Universal Robots PolyScope program: krc_tending.urp

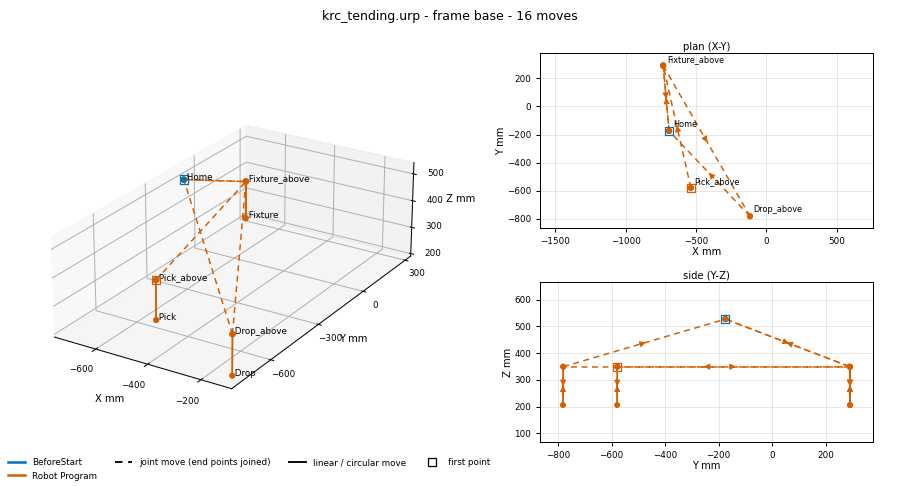
[picture p0: tool path of krc_tending.urp in frame base, 16 of 17 moves have a stored position in this frame; points joined in program order, loops and branches not executed]
Program krc_tending (installation=krc_cell directory=/programs createdIn=5.12.7.1102192 lastSavedIn=5.12.7.1102192 robotSerialNumber=20195299999)
Calibrated DH parameters: a=[0, -0.6127, -0.57155, 0, 0, 0]; d=[0.1807, 0, 0, 0.17415, 0.11985, 0.11655]; alpha=[1.570796, 0, 0, 1.570796, -1.570796, 0]; deltaTheta=[0, 0, 0, 0, 0, 0]
InitVariablesNode
BeforeStart
  'First move: to where the arm already is, so starting the program never moves it on its own'
  start_pose := get_actual_tcp_pose()
  MoveL speed 150 mm/s, acceleration 500 mm/s^2 (useActiveTCP=true optimoveEnabled=false optiMoveSpeed=0.3 optiMoveAcceleration=0.09) feature=Base
    Waypoint Start_pose (Variable): variable=start_pose
  'Every start: clear the handshake, then check it's at home before it moves at all'
  Set ExpressionOutput pin=GP_int_out[5]; expression=10
  Set ExpressionOutput pin=GP_int_out[1]; expression=0
  Set ExpressionOutput pin=GP_int_out[2]; expression=0
  Set ExpressionOutput pin=GP_int_out[3]; expression=0
  Set ExpressionOutput pin=GP_int_out[4]; expression=0
  beat := 0
  home_q := [0.0, -1.57, 1.57, -1.57, -1.57, 0.0]
  q_now := get_actual_joint_positions()
  If norm(q_now[0]-home_q[0])>0.05 or norm(q_now[1]-home_q[1])>0.05 or norm(q_now[2]-home_q[2])>0.05 or norm(q_now[3]-home_q[3])>0.05 or norm(q_now[4]-home_q[4])>0.05 or norm(q_now[5]-home_q[5])>0.05
    'Stopped mid-move last time: moving home from here could hit the fixture or the part, so it doesn't try'
    Set ExpressionOutput pin=GP_int_out[5]; expression=900
    Popup Error (haltProgram=true message=The robot is away from home. Jog it home, then press Start on the panel. inputType=Text)
  Set DigitalOutput pin=tool_out[0]; digitalValue=0
  Wait Sleep waitTime=0.5
  MoveJ speed 57.3 deg/s, acceleration 68.75 deg/s^2 (useActiveTCP=true optimoveEnabled=false optiMoveSpeed=0.3 optiMoveAcceleration=0.09) feature=Base
    Waypoint Home: TCP in base x=-691.676 y=-174.362 z=526.755 mm, rx=2.2206 ry=2.2206 rz=0 rad; joints [0, -89.954, 89.954, -89.954, -89.954, 0] deg; TCP offset x=0 y=0 z=150 mm, rx=0 ry=0 rz=0 rad
Robot Program (runOnlyOnce=false)
  Folder Ready
    'At home, waiting for a command'
    Set ExpressionOutput pin=GP_int_out[5]; expression=100
    Set ExpressionOutput pin=GP_int_out[1]; expression=1
    Wait Condition expression=GP_int_in[1]≟1 or GP_int_in[1]≟2
  Folder Acknowledge
    'Echo the command, and stop being ready while busy'
    cmd := GP_int_in[1]
    Set ExpressionOutput pin=GP_int_out[1]; expression=0
    Set ExpressionOutput pin=GP_int_out[2]; expression=cmd
    ok := True
  If cmd≟1
    'Load: pick a part from the tray, place it in the fixture'
    Set ExpressionOutput pin=GP_int_out[5]; expression=200
    MoveJ speed 57.3 deg/s, acceleration 68.75 deg/s^2 (useActiveTCP=true optimoveEnabled=false optiMoveSpeed=0.3 optiMoveAcceleration=0.09) feature=Base
      Waypoint Pick_above: TCP in base x=-536.89 y=-578.569 z=348.935 mm, rx=2.2208 ry=2.2208 rz=0.001 rad; joints [34.377, -80.214, 97.403, -107.143, -89.954, 34.377] deg
    MoveL speed 150 mm/s, acceleration 500 mm/s^2 (useActiveTCP=true optimoveEnabled=false optiMoveSpeed=0.3 optiMoveAcceleration=0.09) feature=Base
      Waypoint Pick: TCP in base x=-537.712 y=-579.131 z=205.685 mm, rx=2.2208 ry=2.2208 rz=0.001 rad; joints [34.377, -74.485, 105.997, -121.467, -89.954, 34.377] deg
    Set DigitalOutput pin=tool_out[0]; digitalValue=1
    Wait Sleep waitTime=0.5
    MoveL speed 150 mm/s, acceleration 500 mm/s^2 (useActiveTCP=true optimoveEnabled=false optiMoveSpeed=0.3 optiMoveAcceleration=0.09) feature=Base
      Waypoint Pick_above: TCP in base x=-536.89 y=-578.569 z=348.935 mm, rx=2.2208 ry=2.2208 rz=0.001 rad; joints [34.377, -80.214, 97.403, -107.143, -89.954, 34.377] deg
    If tool_out[0]≟False
      'Gripper missed the part'
      ok := False
    Else 
      MoveJ speed 57.3 deg/s, acceleration 68.75 deg/s^2 (useActiveTCP=true optimoveEnabled=false optiMoveSpeed=0.3 optiMoveAcceleration=0.09) feature=Base
        Waypoint Fixture_above: TCP in base x=-733.795 y=290.754 z=348.935 mm, rx=2.2208 ry=2.2208 rz=-0.001 rad; joints [-34.377, -80.214, 97.403, -107.143, -89.954, -34.377] deg
      Set ExpressionOutput pin=GP_int_out[5]; expression=210
      Wait Condition expression=GP_int_in[2]≟1
      MoveL speed 150 mm/s, acceleration 500 mm/s^2 (useActiveTCP=true optimoveEnabled=false optiMoveSpeed=0.3 optiMoveAcceleration=0.09) feature=Base
        Waypoint Fixture: TCP in base x=-734.617 y=291.316 z=205.685 mm, rx=2.2208 ry=2.2208 rz=-0.001 rad; joints [-34.377, -74.485, 105.997, -121.467, -89.954, -34.377] deg
      Set ExpressionOutput pin=GP_int_out[5]; expression=220
      Set DigitalOutput pin=tool_out[0]; digitalValue=0
      Wait Sleep waitTime=0.5
      MoveL speed 150 mm/s, acceleration 500 mm/s^2 (useActiveTCP=true optimoveEnabled=false optiMoveSpeed=0.3 optiMoveAcceleration=0.09) feature=Base
        Waypoint Fixture_above: TCP in base x=-733.795 y=290.754 z=348.935 mm, rx=2.2208 ry=2.2208 rz=-0.001 rad; joints [-34.377, -80.214, 97.403, -107.143, -89.954, -34.377] deg
      MoveJ speed 57.3 deg/s, acceleration 68.75 deg/s^2 (useActiveTCP=true optimoveEnabled=false optiMoveSpeed=0.3 optiMoveAcceleration=0.09) feature=Base
        Waypoint Home: TCP in base x=-691.676 y=-174.362 z=526.755 mm, rx=2.2206 ry=2.2206 rz=0 rad; joints [0, -89.954, 89.954, -89.954, -89.954, 0] deg
  Else 
    'Unload: take the part out of the fixture, drop it'
    Set ExpressionOutput pin=GP_int_out[5]; expression=300
    MoveJ speed 57.3 deg/s, acceleration 68.75 deg/s^2 (useActiveTCP=true optimoveEnabled=false optiMoveSpeed=0.3 optiMoveAcceleration=0.09) feature=Base
      Waypoint Fixture_above: TCP in base x=-733.795 y=290.754 z=348.935 mm, rx=2.2208 ry=2.2208 rz=-0.001 rad; joints [-34.377, -80.214, 97.403, -107.143, -89.954, -34.377] deg
    Wait Condition expression=GP_int_in[2]≟1
    MoveL speed 150 mm/s, acceleration 500 mm/s^2 (useActiveTCP=true optimoveEnabled=false optiMoveSpeed=0.3 optiMoveAcceleration=0.09) feature=Base
      Waypoint Fixture: TCP in base x=-734.617 y=291.316 z=205.685 mm, rx=2.2208 ry=2.2208 rz=-0.001 rad; joints [-34.377, -74.485, 105.997, -121.467, -89.954, -34.377] deg
    Set ExpressionOutput pin=GP_int_out[5]; expression=310
    Set DigitalOutput pin=tool_out[0]; digitalValue=1
    Wait Sleep waitTime=0.5
    MoveL speed 150 mm/s, acceleration 500 mm/s^2 (useActiveTCP=true optimoveEnabled=false optiMoveSpeed=0.3 optiMoveAcceleration=0.09) feature=Base
      Waypoint Fixture_above: TCP in base x=-733.795 y=290.754 z=348.935 mm, rx=2.2208 ry=2.2208 rz=-0.001 rad; joints [-34.377, -80.214, 97.403, -107.143, -89.954, -34.377] deg
    If tool_out[0]≟False
      'Gripper missed the part'
      ok := False
    Else 
      Set ExpressionOutput pin=GP_int_out[5]; expression=320
      MoveJ speed 57.3 deg/s, acceleration 68.75 deg/s^2 (useActiveTCP=true optimoveEnabled=false optiMoveSpeed=0.3 optiMoveAcceleration=0.09) feature=Base
        Waypoint Drop_above: TCP in base x=-116.43 y=-780.664 z=348.935 mm, rx=2.2212 ry=2.2212 rz=0.0016 rad; joints [68.755, -80.214, 97.403, -107.143, -89.954, 68.755] deg
      MoveL speed 150 mm/s, acceleration 500 mm/s^2 (useActiveTCP=true optimoveEnabled=false optiMoveSpeed=0.3 optiMoveAcceleration=0.09) feature=Base
        Waypoint Drop: TCP in base x=-116.791 y=-781.592 z=205.685 mm, rx=2.2212 ry=2.2212 rz=0.0016 rad; joints [68.755, -74.485, 105.997, -121.467, -89.954, 68.755] deg
      Set DigitalOutput pin=tool_out[0]; digitalValue=0
      Wait Sleep waitTime=0.5
      MoveL speed 150 mm/s, acceleration 500 mm/s^2 (useActiveTCP=true optimoveEnabled=false optiMoveSpeed=0.3 optiMoveAcceleration=0.09) feature=Base
        Waypoint Drop_above: TCP in base x=-116.43 y=-780.664 z=348.935 mm, rx=2.2212 ry=2.2212 rz=0.0016 rad; joints [68.755, -80.214, 97.403, -107.143, -89.954, 68.755] deg
      MoveJ speed 57.3 deg/s, acceleration 68.75 deg/s^2 (useActiveTCP=true optimoveEnabled=false optiMoveSpeed=0.3 optiMoveAcceleration=0.09) feature=Base
        Waypoint Home: TCP in base x=-691.676 y=-174.362 z=526.755 mm, rx=2.2206 ry=2.2206 rz=0 rad; joints [0, -89.954, 89.954, -89.954, -89.954, 0] deg
  If ok
    'Done: echo the command'
    Set ExpressionOutput pin=GP_int_out[3]; expression=cmd
  Else 
    'The gripper missed: report fault 1, open, go home'
    Set ExpressionOutput pin=GP_int_out[5]; expression=800
    Set ExpressionOutput pin=GP_int_out[4]; expression=1
    Set DigitalOutput pin=tool_out[0]; digitalValue=0
    Wait Sleep waitTime=0.5
    MoveJ speed 57.3 deg/s, acceleration 68.75 deg/s^2 (useActiveTCP=true optimoveEnabled=false optiMoveSpeed=0.3 optiMoveAcceleration=0.09) feature=Base
      Waypoint Home: TCP in base x=-691.676 y=-174.362 z=526.755 mm, rx=2.2206 ry=2.2206 rz=0 rad; joints [0, -89.954, 89.954, -89.954, -89.954, 0] deg
  Folder Clear
    'Wait for the PLC to drop the command, then clear the handshake'
    Set ExpressionOutput pin=GP_int_out[5]; expression=400
    Wait Condition expression=GP_int_in[1]≟0
    Set ExpressionOutput pin=GP_int_out[2]; expression=0
    Set ExpressionOutput pin=GP_int_out[3]; expression=0
    Set ExpressionOutput pin=GP_int_out[4]; expression=0
Thread 
  'The heartbeat: counts up every 250 ms, as long as this program runs'
  beat := (beat + 1) % 32768
  Set ExpressionOutput pin=GP_int_out[0]; expression=beat
  Wait Sleep waitTime=0.25
